(* IEC 61131-3 sources: moqui-plc/codesys-v4/moqui-plc.fbsdev/moqui.iecapp^/moqui/runtime/component/mantle-hvac/src/main/org/moqui/device, 5 files *)

(* ---- AirDistributionController.fb.st ---- *)
(*
 * AirDistributionController: Logical sequencer for alternating high/low air throw.
 *
 * Implements cumulative timing logic for throw phases:
 * - Time advances only during active operation (operationType = Run AND enable = TRUE).
 * - Counters are frozen (retained) during standby/pause phases.
 * - Implements a Make-Before-Break transition between ducts to prevent overpressure peaks,
 * leveraging the asynchronous handshake mechanism (VAR_IN_OUT) of the underlying Actuator instances.
 *)
FUNCTION_BLOCK AirDistributionController

	VAR_INPUT
	    operationType : OperatingMode := OperatingMode.Init;
	    enable : BOOL; (* Local run permission (e.g., air flow running + air mixing enabled) *)
	    clock1s : BOOL; (* 1-second base clock pulse *)
	END_VAR
	VAR CONSTANT
	    componentName : STRING := 'HVAC_AIR_GROUP';
	END_VAR
	VAR
		(* Logger facade *)
	    logger : LoggerFacade;
	    status : AirDistributionControllerStatus := AirDistributionControllerStatus.Init;
	    cumulatedTimeHigh : UINT := 0;
	    cumulatedTimeLow : UINT := 0;
	    (* Make-before-break: the old damper is disabled only after the new one is enabled *)
	    breakIssued : BOOL;
	END_VAR

	(* Logger facade init *)
	logger.enable := TRUE; logger.loggerName := componentName;

	(* Initialization or reset upon critical Stop *)
	IF operationType = OperatingMode.Init THEN
	    logger(message := 'Init air distribution controller.', level := LogLevel.DEBUG);
	    status := AirDistributionControllerStatus.Init;
	    cumulatedTimeHigh := 0;
	    cumulatedTimeLow := 0;
		ec.dev.highFlowDamperEnableRequest := TRUE;
		ec.dev.highFlowDamperDisableRequest := FALSE;
		ec.dev.lowFlowDamperEnableRequest := FALSE;
		ec.dev.lowFlowDamperDisableRequest := TRUE;
	    RETURN;
	END_IF;

	(* Logic advances ONLY if the system is in Run mode and local enable is active *)
	IF (operationType = OperatingMode.Run) AND enable THEN

	    CASE status OF

	        AirDistributionControllerStatus.Init:
	            (* Startup sequence: defaults to the high throw phase *)
	            ec.dev.highFlowDamperEnableRequest := TRUE;
	 		   	ec.dev.highFlowDamperDisableRequest := FALSE;
	            ec.dev.lowFlowDamperEnableRequest := FALSE;
	 		   	ec.dev.lowFlowDamperDisableRequest := TRUE;
	            logger(message := 'Enter high throw phase.', level := LogLevel.DEBUG);
	            status := AirDistributionControllerStatus.HighPhase;

	        AirDistributionControllerStatus.HighPhase:
	            (* Advance cumulative timer *)
	            IF clock1s THEN
	                cumulatedTimeHigh := cumulatedTimeHigh + 1;
	            END_IF;

	            (* Evaluate switching threshold *)
	            IF ec.dev.setPointTimeHigh > 0 AND cumulatedTimeHigh >= ec.dev.setPointTimeHigh THEN
	                cumulatedTimeHigh := 0;
	                (* Make-Before-Break: first enable the low damper; the high one is disabled in TransitionToLow *)
					ec.dev.lowFlowDamperEnableRequest := TRUE;
					ec.dev.lowFlowDamperDisableRequest := FALSE;
					breakIssued := FALSE;
	                logger(message := 'Transition to low throw.', level := LogLevel.DEBUG);
	                status := AirDistributionControllerStatus.TransitionToLow;
	            END_IF;

	        AirDistributionControllerStatus.TransitionToLow:
	            (* * Monitor the falling edge of the request signals.
	             * The Actuator block internally clears the VAR_IN_OUT variable once
	             * the physical maneuver is completed. This ensures the sequencer
	             * advances only after the hardware has reached its target position.
	             *)
	            IF NOT breakIssued AND NOT ec.dev.lowFlowDamperEnableRequest THEN
	                (* Low damper enabled (make): now disable the high damper (break) *)
					ec.dev.highFlowDamperEnableRequest := FALSE;
					ec.dev.highFlowDamperDisableRequest := TRUE;
					breakIssued := TRUE;
	            ELSIF breakIssued AND NOT ec.dev.highFlowDamperDisableRequest THEN
	                logger(message := 'Enter low throw phase.', level := LogLevel.DEBUG);
	                status := AirDistributionControllerStatus.LowPhase;
	            END_IF;

	        AirDistributionControllerStatus.LowPhase:
	            (* Advance cumulative timer *)
	            IF clock1s THEN
	                cumulatedTimeLow := cumulatedTimeLow + 1;
	            END_IF;

	            (* Evaluate switching threshold *)
	            IF ec.dev.setPointTimeLow > 0 AND cumulatedTimeLow >= ec.dev.setPointTimeLow THEN
	                cumulatedTimeLow := 0;
	                (* Make-Before-Break: first enable the high damper; the low one is disabled in TransitionToHigh *)
					ec.dev.highFlowDamperEnableRequest := TRUE;
					ec.dev.highFlowDamperDisableRequest := FALSE;
					breakIssued := FALSE;
	                logger(message := 'Transition to high throw.', level := LogLevel.DEBUG);
	                status := AirDistributionControllerStatus.TransitionToHigh;
	            END_IF;

	        AirDistributionControllerStatus.TransitionToHigh:
	            (* Wait for hardware positioning confirmation *)
	            IF NOT breakIssued AND NOT ec.dev.highFlowDamperEnableRequest THEN
	                (* High damper enabled (make): now disable the low damper (break) *)
					ec.dev.lowFlowDamperEnableRequest := FALSE;
					ec.dev.lowFlowDamperDisableRequest := TRUE;
					breakIssued := TRUE;
	            ELSIF breakIssued AND NOT ec.dev.lowFlowDamperDisableRequest THEN
	                logger(message := 'Enter high throw phase.', level := LogLevel.DEBUG);
	                status := AirDistributionControllerStatus.HighPhase;
	            END_IF;
	    END_CASE;
	ELSE
	    (* Standby / Pause Condition *)
	    (*
	     * During standby (OperatingMode.Standby OR enable = FALSE), the FB does
	     * not increment any timers. The current status and Request variables are
	     * frozen, maintaining the hardware in its last consolidated stable state.
	     *)
	    ;
	END_IF;
	END_FUNCTION_BLOCK

(* ---- DeviceDiagnostics.fb.st ---- *)
(* Device diagnostics *)
FUNCTION_BLOCK DeviceDiagnostics

	VAR_INPUT
		operationType : OperatingMode := OperatingMode.Run;
	END_VAR
	VAR_OUTPUT
		error : BOOL;
	END_VAR

	error := TRUE;

	(* Signal management engine *)
	(*
	 * Prepare a fresh scan (clears the accumulated output action).
	 * Then process each device signal in priority order.
	 * ImmediateStop -> faultRequest := TRUE -> Main enters Fault state.
	 *)
	ec.dev.signalMgmt(operationType := SignalMgmtOperatingMode.Prepare);
	ec.dev.signalMgmt.operationType := SignalMgmtOperatingMode.Process;

	(* Device faults *)
	ec.dev.signalMgmt(
		loggerName := ec.dev.ahuFan.loggerName,
		code := 16#0001,
		category := SignalCategory.Alarm,
		resetPol := ResetPolicy.UnconditionedReset,
		activationCondition := ec.dev.ahuFan.invalidConfig,
		outputAction := SignalOutputAction.ImmediateStop);
	ec.dev.signalMgmt(
		loggerName := ec.dev.airFlow.loggerName,
		code := 16#0002,
		category := SignalCategory.Alarm,
		resetPol := ResetPolicy.UnconditionedReset,
		activationCondition := ec.dev.airFlow.fault,
		outputAction := SignalOutputAction.ImmediateStop);
	ec.dev.signalMgmt(
		loggerName := ec.dev.coldGlycolPump.loggerName,
		code := 16#0003,
		category := SignalCategory.Alarm,
		resetPol := ResetPolicy.UnconditionedReset,
		activationCondition := ec.dev.coldGlycolPump.fault,
		outputAction := SignalOutputAction.ImmediateStop);
	ec.dev.signalMgmt(
		loggerName := ec.dev.coldGlycolValve.loggerName,
		code := 16#0004,
		category := SignalCategory.Alarm,
		resetPol := ResetPolicy.UnconditionedReset,
		activationCondition := ec.dev.coldGlycolValve.invalidConfig,
		outputAction := SignalOutputAction.ImmediateStop);
	ec.dev.signalMgmt(
		loggerName := ec.dev.hotGlycolPump.loggerName,
		code := 16#0005,
		category := SignalCategory.Alarm,
		resetPol := ResetPolicy.UnconditionedReset,
		activationCondition := ec.dev.hotGlycolPump.fault,
		outputAction := SignalOutputAction.ImmediateStop);
	ec.dev.signalMgmt(
		loggerName := ec.dev.hotGlycolValve.loggerName,
		code := 16#0006,
		category := SignalCategory.Alarm,
		resetPol := ResetPolicy.UnconditionedReset,
		activationCondition := ec.dev.hotGlycolValve.invalidConfig,
		outputAction := SignalOutputAction.ImmediateStop);
	ec.dev.signalMgmt(
		loggerName := ec.dev.highFlowDamper.loggerName,
		code := 16#0007,
		category := SignalCategory.Alarm,
		resetPol := ResetPolicy.UnconditionedReset,
		activationCondition := ec.dev.highFlowDamper.fault,
		outputAction := SignalOutputAction.ImmediateStop);
	ec.dev.signalMgmt(
		loggerName := ec.dev.lowFlowDamper.loggerName,
		code := 16#0008,
		category := SignalCategory.Alarm,
		resetPol := ResetPolicy.UnconditionedReset,
		activationCondition := ec.dev.lowFlowDamper.fault,
		outputAction := SignalOutputAction.ImmediateStop);

	(*
	 * Duct safety alarms - supply-air temperature limits (ImmediateStop).
	 * Air that is too hot or too cold entering the curing room can damage
	 * or contaminate the product. These alarms are always evaluated
	 * regardless of the current FSM state.
	 *)
	ec.dev.signalMgmt(
		loggerName := 'HVAC_DEMO_PLC',
		code := 16#0010,
		category := SignalCategory.Alarm,
		resetPol := ResetPolicy.UnconditionedReset,
		activationCondition := ec.dev.ductTempOverMax,
		outputAction := SignalOutputAction.ImmediateStop);
	ec.dev.signalMgmt(
		loggerName := 'HVAC_DEMO_PLC',
		code := 16#0011,
		category := SignalCategory.Alarm,
		resetPol := ResetPolicy.UnconditionedReset,
		activationCondition := ec.dev.ductTempUnderMin,
		outputAction := SignalOutputAction.ImmediateStop);

	(* Duct RH - Warning only (condensation risk, does not stop the machine) *)
	ec.dev.signalMgmt(
		loggerName := 'HVAC_DEMO_PLC',
		code := 16#0012,
		category := SignalCategory.Warning,
		resetPol := ResetPolicy.UnconditionedReset,
		activationCondition := ec.dev.ductRhOverMax,
		outputAction := SignalOutputAction.None);

	error := FALSE;
	END_FUNCTION_BLOCK

(* ---- DeviceManager.fb.st ---- *)
(* Hardware Abstraction Layer (HAL) orchestrator.
 *
 * Drives all physical device FBs once per scan.
 * Main component sets the enable/disable request flags; DeviceManager wires them
 * to the individual Actuator / ProcessPid FBs.
 *
 * Call order within the PLC task:
 *   InputSignalUpdate (updates feedback signals from field)
 *   Main (FSM + MainRuleEngine -> sets request flags)
 *   DeviceManager (this block - drives device FBs)
 *   OutputSignalUpdate (maps device outputs to physical terminals)
 *
 * Handshake note (Actuator FBs):
 *   enableRequest / disableRequest are VAR_IN_OUT.  The Actuator FB clears
 *   the flag as its acknowledgment.  Main.pou re-asserts the flag each scan
 *   from dev.xxxEnableRequest, so the handshake is level-triggered.
 *
 * ProcessPid note (ahuFan):
 *   ProcessPid uses a plain BOOL 'enable' input - no VAR_IN_OUT handshake.
 *   Setting enable := FALSE ramps the output to 0 and disables the controller.
 *)
FUNCTION_BLOCK DeviceManager

	VAR_INPUT
		operationType : OperatingMode := OperatingMode.Run;
	END_VAR

	(* Cold glycol group *)
	(*
	 * Pump is started first via the request/ack handshake.
	 * The valve follows the pump state, not the request: the pump clears
	 * coldGroupEnableRequest as its acknowledgment, so the request is FALSE
	 * exactly while the group is running (enable := FALSE freezes the output at 0).
	 *)
	ec.dev.coldGlycolPump(
		operationType := operationType,
		clock := ec.clks.clock100ms,
		enableRequest := ec.dev.coldGroupEnableRequest,
		disableRequest := ec.dev.coldGroupDisableRequest);

	(* Reverse acting: cooling opens the valve when the temperature is above the setpoint *)
	ec.dev.coldGlycolValve(
		enable := ec.dev.coldGlycolPump.isEnabled,
		deviationInversion := TRUE,
		feedback := ec.dev.tempFeedback,
		setpoint := ec.dev.tempSetpoint,
		clock := ec.clks.clock100ms);

	(* Hot glycol group *)
	ec.dev.hotGlycolPump(
		operationType := operationType,
		clock := ec.clks.clock100ms,
		enableRequest := ec.dev.hotGroupEnableRequest,
		disableRequest := ec.dev.hotGroupDisableRequest);

	ec.dev.hotGlycolValve(
		enable := ec.dev.hotGlycolPump.isEnabled,
		feedback := ec.dev.tempFeedback,
		setpoint := ec.dev.tempSetpoint,
		clock := ec.clks.clock100ms);

	(* AHU fan *)
	(*
	 * enable := FALSE ramps down the drive and disables the PID output.
	 * Speed setpoint (ahuFanSpeedSetpoint) and the PID tuning parameters
	 * (gain, integrationTime, etc.) are mapped from the device config (recipe).
	 * ahuFanSpeedFeedback is wired from InputSignalUpdate (drive feedback word).
	 *)
	ec.dev.ahuFan(
		enable := ec.dev.ahuFanEnableRequest,
		setpoint := ec.dev.ahuFanSpeedSetpoint,
		feedback := ec.dev.ahuFanSpeedFeedback,
		clock := ec.clks.clock100ms);

	(* Air flow distributor (drive) *)
	(*
	 * Treated as Actuator with an additional speed reference.
	 * ref = distribution setpoint (0-100 %) from device config (recipe)/RuleEngine.
	 * feedback = drive speed feedback from InputSignalUpdate.
	 * The drive alternates supply air between left and right ducts
	 * according to the ref timing programmed on the drive itself;
	 * the PLC only starts / stops it and adjusts the reference level.
	 *)
	ec.dev.airFlow(
		operationType := operationType,
		clock := ec.clks.clock100ms,
		enableRequest := ec.dev.airFlowEnableRequest,
		disableRequest := ec.dev.airFlowDisableRequest,
		ref := ec.dev.airFlowRef,
		feedback := ec.dev.airFlowSpeedFeedback);

	(* High Flow Damper *)
	(* Requests are generated by AirDistributionController when air mixing is enabled. *)
	ec.dev.highFlowDamper(
		operationType := operationType,
		clock := ec.clks.clock100ms,
		enableRequest := ec.dev.highFlowDamperEnableRequest,
		disableRequest := ec.dev.highFlowDamperDisableRequest);

	(* Low Flow Damper *)
	(* Requests are generated by AirDistributionController when air mixing is enabled. *)
	ec.dev.lowFlowDamper(
		operationType := operationType,
		clock := ec.clks.clock100ms,
		enableRequest := ec.dev.lowFlowDamperEnableRequest,
		disableRequest := ec.dev.lowFlowDamperDisableRequest);
	END_FUNCTION_BLOCK

(* ---- InputSignalUpdate.fb.st ---- *)
(*
 * Input signal acquisition and pre-processing unit.
 * Map physical input terminals/signals to their logical parameters, performing pre-processing (e.g.: signal filtering) if necessary.
 *)
FUNCTION_BLOCK InputSignalUpdate

	VAR_INPUT
		operationType : OperatingMode;
	END_VAR
	VAR
		(* Logger facade *)
		logger : LoggerFacade;
	END_VAR

	(* Logger facade init *)
	logger.enable := TRUE; logger.loggerName := MoquiConf.applicationDeviceId;

	logger(message := 'Input signals acquisition and pre-processing.', level := LogLevel.DEBUG);

	(*
		Physical to logical terminals mapping example:

		IF operationType = OperatingMode.Init THEN
			(* Special processing for the init phase, if needed, such as the restart phase after a blackout. *)
			(* etc. *)
		ELSIF operationType = OperatingMode.Run THEN
			(* Example mapping of 32 bits and 64 bits analog signals *)
			dev.speedFeedback := doubleWordToReal(wordArray := io.speedFeedbackSignal);
			dev.speedFeedback := longWordToLongReal(wordArray := io.speedFeedbackSignal);
			(* Reverse logic *)
			dev.coldGlycolValve.disabledSensor := NOT io.coldGlycolValveSignalingContact;

			outletColdGlycolTemp := TO_REAL(outletColdGlycolTempSignal);
			(* Analog input processing (scaling, limiting, etc. *)
			dev.tempFeedback := processAnalogInput(io.tempFeedbackSignal, 0, 27000, dev.tempMin, dev.tempMax, -20, 70, 0);
			(* Analog input exponential (1-pole) filtering *)
			expFilter(input := io.coldGlycolTempSignal, t:= 3, start := TRUE, timeElapsed => timeElapsed);
			IF timeElapsed >= 3 THEN dev.outletColdGlycolTemp := expFilter.output; END_IF;
			(* Digital input processing (filtering, debouncing, reverse logic, etc. *)
			digitalFilter(signal := io.airFlowEnabledSensor, enableDelay := T#10MS, disableDelay := T#15MS);
			dev.airFlow.enabledSensor := digitalFilter.delayedSignal;
			(* Drive status word, feedbacks, etc. mapping *)
			processDriveCyclicInData(model := DriveModel.ABBACH580, statusWord := io.compressorStatusWord,
				enabledSensor => dev.compressor.enabledSensor, disabledSensor => dev.compressor.disabledSensor,
				externalFault => dev.compressorExternalFault);
			dev.speedFeedback := TO_REAL(speedFeedbackSignal);
			dev.coldGlycolPump.enabledSensor := io.coldGlycolPumpAuxContact;
			dev.coldGlycolPump.disabledSensor := NOT io.coldGlycolPumpAuxContact;
			dev.coldGlycolPumpThermistors := io.coldGlycolPumpThermistors;
			dev.coldGlycolFlowSwitch := io.coldGlycolFlowSwitch;
			dev.coldGlycolPumpPowerSupplyFault := NOT io.coldGlycolPumpShuntTrip;
			dev.coldGlycolCircPumpExternalFault := io.coldGlycolPumpShuntTrip OR io.coldGlycolPumpThermistors
				OR io.coldGlycolFlowSwitch;
			...

		END_IF;

		(*
		 * Configure and call the logger facade to log signals where needed.
		 *     logger(payloadType := LogPayloadType.Numeric, numericValue := dev.speedRef, level := LogLevel.DEBUG);
		 *     logger(payloadType := LogPayloadType.Numeric, numericValue := dev.outletColdGlycolTemp, level := LogLevel.DEBUG);
		 *     (* etc. *)
		 *)
	*)
	END_FUNCTION_BLOCK

(* ---- OutputSignalUpdate.fb.st ---- *)
(*
 * Output signals processing (e.g.: debouncing filter) and actuation unit.
 * Map logical output parameters on their physical counterpart, performing processing if necessary.
 *)
FUNCTION_BLOCK OutputSignalUpdate

	VAR_INPUT
		operationType : OperatingMode;
	END_VAR
	VAR
		(* Logger facade *)
		logger : LoggerFacade;
	END_VAR

	(* Logger facade init *)
	logger.enable := TRUE; logger.loggerName := MoquiConf.applicationDeviceId;

	logger(message := 'Output signals processing and actuation.', level := LogLevel.DEBUG);

	(*
		Logical to physical terminals mapping example:

		IF operationType = OperatingMode.Init THEN
			(* Special processing for the init phase, if needed, such as the restart phase after a blackout. *)
			(* etc. *)
		ELSIF operationType = OperatingMode.Run THEN
			(* For continuous speed values mapping ... *)
			(* Example mapping of a word analog signal *)
			io.speedRefSignal := TO_WORD(dev.speedRef);
			(* Example mapping of a 32-bit analog signal *)
			io.speedRefSignal := realToWordArray(dev.speedRef);
			(* Example mapping of a 64-bit analog signal *)
			io.speedRefSignal := longRealToWordArray(dev.speedRef);
			io.coldGlycolTempSignal := TO_WORD(dev.inletColdGlycolTemp);
			(* Scaling and limiting example *)
			processAnalogOutput(dev.tempSetpoint, 4, 20, dev..tempMin,
				dev.tempMax, 0, 1, 0, wordAnalogOutput => io.tempSetpointSignal);
			(* Drive control word and reference mapping *)
			processDriveCyclicOutData(DriveModel.ABBACH580, dev.compressor.enable, reset := FALSE,
				controlWord => io.compressorControlWord);
			(* Reverse logic *)
			io.condenserFanEnableContactor := NOT condenserFan.enable;
			io.coldGlycolPumpContactor := dev.coldGlycolPump.enable;
			io.coldGlycolPumpContactor := NOT dev.coldGlycolPump.disable;
			io.faultLight := coldGlycolPump.fault;
			...
		END_IF;

		(*
		 * Configure and call the logger facade to log signals where needed.
		 *     logger(payloadType := LogPayloadType.Numeric, numericValue := io.speedRefSignal, level := LogLevel.DEBUG);
		 *     logger(payloadType := LogPayloadType.Numeric, numericValue := io.coldGlycolTempSignal, level := LogLevel.DEBUG);
		 *     logger(payloadType := LogPayloadType.Enum, enumValue := io.controlWord, level := LogLevel.DEBUG);
		 *     (* etc. *)
		 *)
	*)
	END_FUNCTION_BLOCK
